SUBAPPLICATION Uebung_011d_GcfFunc_AX (* Numeric Value Input I1 Durchschleifen auf N3 (Offset/Scale Effekt) *)
  (* Standard: 61499-2; Description: Copyright (c) 2023 Meisterschulen am Ostbahnhof This program and the accompanying materials are made available under the terms of the Eclipse Public License 2.0 which is available at https://www.eclipse.org/legal/epl-2.0/ SPDX-License-Identifier: EPL-2.0 *)
  (* Version 1.0, 2026-04-14, Franz Höpfinger, Meisterschulen am Ostbahnhof, initial API and implementation and/or initial documentation *)
  PACKAGE Meins::GcfFunctionCall;
  IMPORT Meins::GcfFunctionCall::const::FuncConst::DOUBLE_VALUE;
  IMPORT Uebungen::const::UT::DefaultPool_Numeric::OutputNumber_N3_N;
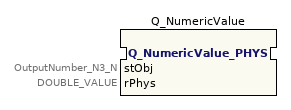
  FBS
    Q_NumericValue : isobus::UT::Q::Q_NumericValue_PHYS(stObj := OutputNumber_N3_N, rPhys := DOUBLE_VALUE);
  END_FBS
END_SUBAPPLICATION
